// TIA Portal V21 export
Screen "Pump"  NonexNone, Number=2
  ScreenLayer 
    TextField "SpeedLabel" at 20,40 size 160x30  Text="<body><p>Pump speed</p></body>"
    IOField "SpeedValue" at 200,40 size 120x30
